{attribute 'qualified_only'}
{attribute 'strict'}
TYPE EJECT_ENUM :
(
	YES := 0,
	NO_2_START := 1,
	NO_1_START := 2
)UDINT;
END_TYPE

(* stored: Version 1.1.0.1, ProductVersion 3.1.4024.12
   DUT EJECT_ENUM: Id {399122cf-8424-444c-b905-9341d13cde4e} *)
